  def log_weight():
  	socket_open(SERVER_IP,SERVER_PORT)
  	socket_send_string("LOG_WEIGHT")
  	sleep(0.5)
  	socket_close()
  end

  def send_target_info():
  	socket_open(SERVER_IP,SERVER_PORT)
  	socket_send_string("SET_TARGET:" + to_str(target_weight))
  	sleep(0.2)
  	socket_close()
  end
  def send_powder_info():
  	socket_open(SERVER_IP,SERVER_PORT)
  	socket_send_string("SET_POWDER:" + Pow_name)
  	sleep(0.2)
  	socket_close()
  end
  def send_spatula_info():
  	socket_open(SERVER_IP,SERVER_PORT)
  	socket_send_string("SET_SPATULA:" + spatula)
  	#sleep(1)

  	#local fl = socket_read_ascii_float(4)
    	#socket_close()

    	#global s_depth = fl[1]
    	#global s_length = fl[2]
   	#global s_volume = fl[3]
   	#global ry_theta  = fl[4]
  	sleep(0.2)

  end

  def send_level_info():
  	socket_open(SERVER_IP,SERVER_PORT)
  	socket_send_string("SET_LEVEL:" + to_str(level))
  	sleep(0.2)
  	socket_close()
  end

  def get_cont_weight():
    socket_open(SERVER_IP, SERVER_PORT)
    #rq_open_and_wait()
    cmd = "GET_CONT_WEIGHT"
    socket_send_string(cmd)
    sync()
    sleep(0.5)
    receiveFromSer = socket_read_ascii_float(1)
    socket_close()
    return receiveFromSer[1]
  end

  $ 22 "BeforeStarts"
  $ 23 "uLM"
  $ 24 "CMD_Stop≔ False "
  global CMD_Stop=  False
  $ 25 "CMD_Abort≔ False "
  global CMD_Abort=  False
  $ 26 "CMD_Clear≔ False "
  global CMD_Clear=  False
  $ 27 "STATE≔1"
  global STATE=1
  $ 28 "STATE_Info≔''"
  global STATE_Info=""
  $ 29 "ARM_Referenced≔ False "
  global ARM_Referenced=  False
  $ 30 "zero_ftsensor()"
  zero_ftsensor()
  $ 31 "poses init"
  $ 32 "PSE_A≔p[0,0,0,0,0,0]"
  global PSE_A=p[0,0,0,0,0,0]
  $ 33 "PSE_A_H≔p[0,0,0,0,0,0]"
  global PSE_A_H=p[0,0,0,0,0,0]
  $ 34 "PSE_R≔p[0,0,0,0,0,0]"
  global PSE_R=p[0,0,0,0,0,0]
  $ 35 "PSE_R_H≔p[0,0,0,0,0,0]"
  global PSE_R_H=p[0,0,0,0,0,0]
  $ 36 "PSE_T≔p[0,0,0,0,0,0]"
  global PSE_T=p[0,0,0,0,0,0]
  $ 37 "PSE_T_H≔p[0,0,0,0,0,0]"
  global PSE_T_H=p[0,0,0,0,0,0]
  $ 38 "PSE_C_E≔p[0,0,0,0,0,0]"
  global PSE_C_E=p[0,0,0,0,0,0]
  $ 39 "PSE_C_H≔p[0,0,0,0,0,0]"
  global PSE_C_H=p[0,0,0,0,0,0]
  $ 40 "PSE_C_S≔p[0,0,0,0,0,0]"
  global PSE_C_S=p[0,0,0,0,0,0]
  $ 41 "init_home_by_cartesian_pose(p[0,-0.400,0.300,0,0,0])"
  init_home_by_cartesian_pose(p[0,-0.400,0.300,0,0,0])
  $ 42 "Clearing"
  $ 43 "reset_error()"
  reset_error()
  $ 44 "reset_warning()"
  reset_warning()
  $ 45 "uGo"
  $ 47 "ugo_init( True ,'http://192.168.12.120:10001')"
  ugo_init(  True  ,"http://192.168.12.120:10001")
  $ 48 "ugo_update_outputs()"
  ugo_update_outputs()
  $ 49 "App"
  $ 50 "'ADD APPLICATION SPECIFIC COMMANDS'"
  # 'ADD APPLICATION SPECIFIC COMMANDS'
  $ 51 "Tools"
  $ 52 "OBJ_Picked≔gripper_has_object()"
  global OBJ_Picked=gripper_has_object()
  $ 53 "If OBJ_Picked"
  if (OBJ_Picked):
    # begin: URCap Program Node
    #   Source: Robotiq_Grippers, 3.17.0.105337, Robotiq Inc.
    #   Type: Gripper Activate
    $ 54 "Gripper Activate"

    kill rq_gripper_communication_thread
    rq_gripper_communication_thread_started = False
    rq_close_gripper_socket("1")
    rq_close_gripper_socket("2")
    rq_close_gripper_socket("3")
    rq_close_gripper_socket("4")

    rq_init_comm_if_connected(9, "1")
    rq_init_comm_if_connected(2, "2")
    rq_init_comm_if_connected(3, "3")
    rq_init_comm_if_connected(4, "4")
    rq_print_connected_grippers()
    rq_gripper_communication_thread = run rq_gripper_communication()

    while(not rq_gripper_communication_thread_started):
        sleep(0.008)
    end

    rq_set_max_current_for_all_grippers()

    reset_and_activate = False

    rq_activate_all_grippers(False)
    # end: URCap Program Node
  else:
    $ 55 "Else" "noBreak"
    # begin: URCap Program Node
    #   Source: Robotiq_Grippers, 3.17.0.105337, Robotiq Inc.
    #   Type: Gripper Activate
    $ 56 "Gripper Reset and Activate"

    kill rq_gripper_communication_thread
    rq_gripper_communication_thread_started = False
    rq_close_gripper_socket("1")
    rq_close_gripper_socket("2")
    rq_close_gripper_socket("3")
    rq_close_gripper_socket("4")

    rq_init_comm_if_connected(9, "1")
    rq_init_comm_if_connected(2, "2")
    rq_init_comm_if_connected(3, "3")
    rq_init_comm_if_connected(4, "4")
    rq_print_connected_grippers()
    rq_gripper_communication_thread = run rq_gripper_communication()

    while(not rq_gripper_communication_thread_started):
        sleep(0.008)
    end

    rq_set_max_current_for_all_grippers()

    reset_and_activate = True

    rq_activate_all_grippers(True)
    # end: URCap Program Node
  end
  $ 57 "zero_ftsensor()"
  zero_ftsensor()
  $ 58 "EXTT"
  $ 59 "Set GRP_3F_Enable=Off"
  set_standard_digital_out(4, False)
  $ 60 "Set BarcodeTrigger=Off"
  set_standard_digital_out(6, False)
  $ 61 "Set GRP_3F_Decap=Off"
  set_standard_digital_out(3, False)
  $ 62 "Set GRP_3F_Cap=Off"
  set_standard_digital_out(2, False)
  $ 63 "Set GRP_3F_Open=Off"
  set_standard_digital_out(5, False)
  $ 64 "PSE_T≔get_tool_free_pose(dir=[0,0,0.150], move_in_base_frame=True)"
  global PSE_T=get_tool_free_pose(dir=[0,0,0.150], move_in_base_frame=True)
  $ 65 "If is_reachable(Base_const, [PSE_T])"
  if (is_reachable(p[0.0,0.0,0.0,0.0,0.0,0.0], [PSE_T])):
    $ 66 "MoveL"
    $ 67 "PSE_T" "breakAfter"
    movel(PSE_T, a=1.2, v=0.15)
  end
  $ 68 "powder dispensing variable init"
  $ 69 "Start_thread≔ False "
  global Start_thread=  False
  $ 70 "vib_thread≔ False "
  global vib_thread=  False
  $ 71 "w_full_thread≔ False "
  global w_full_thread=  False
  $ 72 "d_cc≔0.07"
  global d_cc=0.07
  $ 73 "kp≔0.0035"
  global kp=0.0035
  $ 74 "ki≔0.0001"
  global ki=0.0001
  $ 75 "kd≔0.003"
  global kd=0.003
  $ 76 "dt≔0.2"
  global dt=0.2
  $ 77 "Integral_error≔0"
  global Integral_error=0
  $ 78 "current_error≔0"
  global current_error=0
  $ 79 "previous_error≔0"
  global previous_error=0
  $ 80 "tilt_increment≔0"
  global tilt_increment=0
  $ 81 "tilt_angle≔0"
  global tilt_angle=0
  $ 82 "diff≔0"
  global diff=0
  $ 83 "tilt_to_home()"
  tilt_to_home()
  $ 84 "switch_spat_M≔ True "
  global switch_spat_M=  True
  $ 85 "switch_spat_S≔ True "
  global switch_spat_S=  True
  $ 86 "switch_spat_F_M≔ True "
  global switch_spat_F_M=  True
  $ 87 "switch_spat_F_S≔ True "
  global switch_spat_F_S=  True
  $ 88 "last_scale≔0"
  global last_scale=0
  $ 817 "Thread_1"
  thread Thread_1():
    while (True):
      $ 818 "If Start_thread≟ True "
      if (Start_thread ==   True  ):
        $ 819 "weight_value≔get_weight()"
        global weight_value=get_weight()
        $ 820 "diff≔target_weight-weight_value"
        global diff=target_weight-weight_value
        $ 821 "Wait: 0.2"
        sleep(0.2)
        $ 822 "sync()"
        sync()
      end
      $ 823 "sync()"
      sync()
    end
  end
  threadId_Thread_1 = run Thread_1()
  $ 824 "Thread_2"
  thread Thread_2():
    while (True):
      $ 825 "Loop vib_thread≟ True "
      thread Thread_while_825():
        while (True):
          $ 826 "diff≔target_weight-weight_value"
          global diff=target_weight-weight_value
          $ 827 "If diff>0.02 and spatula≠'spatula_flat_S' "
          global thread_flag_827=0
          thread Thread_if_827():
            $ 829 "Set AO[0]=4.0"
            set_standard_analog_out(0, 0.4)
            thread_flag_827 = 1
          end
          if (diff>0.02  and  spatula != "spatula_flat_S" ):
            global thread_handler_827=run Thread_if_827()
            while (thread_flag_827 == 0):
              if not(diff>0.02  and  spatula != "spatula_flat_S" ):
                kill thread_handler_827
                thread_flag_827 = 2
              else:
                sync()
              end
            end
          else:
            thread_flag_827 = 2
          end
          if (thread_flag_827 == 2):
            $ 830 "ElseIf diff>0.02 and spatula≟'spatula_flat_S'"
            if (diff>0.02 and spatula == "spatula_flat_S"):
              $ 831 "vibration_3()"
              vibration_3()
            else:
              $ 832 "ElseIf diff≤0.03"
              global thread_flag_832=0
              thread Thread_if_832():
                $ 833 "vibration_2()"
                vibration_2()
                thread_flag_832 = 1
              end
              if (diff <= 0.03):
                global thread_handler_832=run Thread_if_832()
                while (thread_flag_832 == 0):
                  if not(diff <= 0.03):
                    kill thread_handler_832
                    thread_flag_832 = 2
                  else:
                    sync()
                  end
                end
              else:
                thread_flag_832 = 2
              end
              if (thread_flag_832 == 2):
                $ 834 "Else" "noBreak"
                $ 835 "Set AO[0]=0.0"
                set_standard_analog_out(0, 0.0)
              end
            end
          end
        end
      end
      if (vib_thread ==   True  ):
        global thread_handler_825=run Thread_while_825()
        while (vib_thread ==   True  ):
          sync()
        end
        kill thread_handler_825
      end
      $ 836 "sync()"
      sync()
    end
  end
  threadId_Thread_2 = run Thread_2()
  $ 837 "Thread_3"
  thread Thread_3():
    while (True):
      $ 838 "If w_full_thread≟ True "
      if (w_full_thread ==   True  ):
        $ 839 "aa_weight_cont≔get_cont_weight()"
        global aa_weight_cont=get_cont_weight()
        $ 840 "Wait: 0.2"
        sleep(0.2)
        $ 841 "sync()"
        sync()
      end
      $ 842 "sync()"
      sync()
    end
  end
  threadId_Thread_3 = run Thread_3()
  while (True):
    $ 89 "Robot Program"
    $ 90 "MAIN"
    $ 91 "command_manager(external_control='uGO', cond_suspend=(ITM_Manipulated and AMR_AtTarget and AMR_Charging and AMR_Battery<40), cond_unsuspend=(AMR_Battery≟60))"
    command_manager(external_control="uGO", cond_suspend=(ITM_Manipulated  and  AMR_AtTarget  and  AMR_Charging  and  AMR_Battery<40), cond_unsuspend=(AMR_Battery == 60))
    $ 92 "log_state(STATE_Info)"
    log_state(STATE_Info)
    $ 93 "Switch STATE"
    switch_1 = STATE
    $ 94 "Case 1"
    if (1 == switch_1):
      $ 95 "Stopping"
      $ 96 "STATE_Info≔'Stopping'"
      global STATE_Info="Stopping"
      $ 97 "end_freedrive_mode()"
      end_freedrive_mode()
      $ 98 "Set"
      set_tcp(p[0.0,0.0,0.161,3.1415,0.0,0.0])
      $ 99 "PSE_T≔get_tool_free_pose(dir=[0,0,0.150], move_in_base_frame=True)"
      global PSE_T=get_tool_free_pose(dir=[0,0,0.150], move_in_base_frame=True)
      $ 100 "If is_reachable(Base_const, [PSE_T])"
      if (is_reachable(p[0.0,0.0,0.0,0.0,0.0,0.0], [PSE_T])):
        $ 101 "MoveL"
        $ 102 "PSE_T" "breakAfter"
        movel(PSE_T, a=1.2, v=0.15)
      end
      $ 103 "do_transition(keep_rxry=OBJ_Picked, r=0)"
      do_transition(keep_rxry=OBJ_Picked, r=0)
      $ 112 "Call Sub_AMR_MiR_V3"
      Sub_AMR_MiR_V3()
      $ 113 "If stopping() and AMR_Done"
      if (stopping()  and  AMR_Done):
        $ 114 "STATE≔2"
        global STATE=2
        $ 115 "ugo_update_outputs()"
        ugo_update_outputs()
      end
    elif (2 == switch_1):
      $ 116 "Case 2"
      $ 117 "Stopped"
      $ 118 "STATE_Info≔'Stopped'"
      global STATE_Info="Stopped"
      $ 119 "Call Sub_AMR_MiR_V3"
      Sub_AMR_MiR_V3()
      $ 120 "If CMD_Reset  or PB_Start"
      if (CMD_Reset   or  get_standard_digital_in(0)):
        $ 121 "STATE≔3"
        global STATE=3
        $ 122 "ugo_update_outputs()"
        ugo_update_outputs()
      end
    elif (3 == switch_1):
      $ 123 "Case 3"
      $ 124 " Resetting"
      $ 125 "STATE_Info≔'Resetting'"
      global STATE_Info="Resetting"
      $ 126 "uML"
      $ 127 "reset_error()"
      reset_error()
      $ 128 "reset_warning()"
      reset_warning()
      $ 129 "PROCESS_Step≔0"
      global PROCESS_Step=0
      $ 130 "PROCESS_Info≔''"
      global PROCESS_Info=""
      $ 131 "ARM_Referenced≔ False "
      global ARM_Referenced=  False
      $ 132 "WRK_Done≔ False "
      global WRK_Done=  False
      $ 133 "ITM_Prepared≔ False "
      global ITM_Prepared=  False
      $ 134 "ITM_Manipulated≔ False "
      global ITM_Manipulated=  False
      $ 135 "STP≔0"
      global STP=0
      $ 136 "Action≔0"
      global Action=0
      $ 137 "Action_Info≔''"
      global Action_Info=""
      $ 138 "ITM_ID≔0"
      global ITM_ID=0
      $ 139 "JIG≔0"
      global JIG=0
      $ 140 "JIG_Slot≔0"
      global JIG_Slot=0
      $ 141 "Task_info≔''"
      global Task_info=""
      $ 142 "Set"
      set_tcp(p[0.0,0.0,0.161,3.1415,0.0,0.0])
      $ 143 "App"
      $ 144 "'ADD APPLICATION SPECIFIC COMMANDS'"
      # 'ADD APPLICATION SPECIFIC COMMANDS'
      $ 145 "OBJ_Type≔0"
      global OBJ_Type=0
      $ 146 "OBJ_Nbr≔0"
      global OBJ_Nbr=0
      $ 147 "If CNT_Rack_Output≥50"
      if (CNT_Rack_Output >= 50):
        $ 148 "CNT_Rack_Output≔0"
        global CNT_Rack_Output=0
      end
      $ 149 "TASK≔struct(ID=0, NAVI=struct(target=0, footprint=0, protectiveOff=0, dock=0), WORK=struct(ITM_ID_Src=0, JIG_ID_Src=0, OBJ_Nbr_Src=0, ACT_Src=0, ITM_ID_Tgt=0, JIG_ID_Tgt=0, OBJ_Nbr_Tgt=0, ACT_Tgt=0, OBJ_Type=0))"
      global TASK=struct(ID=0, NAVI=struct(target=0, footprint=0, protectiveOff=0, dock=0), WORK=struct(ITM_ID_Src=0, JIG_ID_Src=0, OBJ_Nbr_Src=0, ACT_Src=0, ITM_ID_Tgt=0, JIG_ID_Tgt=0, OBJ_Nbr_Tgt=0, ACT_Tgt=0, OBJ_Type=0))
      $ 150 "Call Sub_AMR_MiR_V3"
      Sub_AMR_MiR_V3()
      $ 151 "If resetting() and AMR_Done"
      if (resetting()  and  AMR_Done):
        $ 152 "STATE≔4"
        global STATE=4
        $ 153 "ugo_update_outputs()"
        ugo_update_outputs()
      end
    elif (4 == switch_1):
      $ 154 "Case 4"
      $ 155 "Idle"
      $ 156 "STATE_Info≔'Idle'"
      global STATE_Info="Idle"
      $ 157 "If CMD_Start"
      if (CMD_Start):
        $ 158 "STATE≔5"
        global STATE=5
        $ 159 "ugo_update_outputs()"
        ugo_update_outputs()
      end
    elif (5 == switch_1):
      $ 160 "Case 5"
      $ 161 "Starting"
      $ 162 "STATE_Info≔'Starting'"
      global STATE_Info="Starting"
      $ 163 "'ADD COMMANDS WHAT TO START WITH'"
      # 'ADD COMMANDS WHAT TO START WITH'
      $ 164 "Call Sub_AMR_MiR_V3"
      Sub_AMR_MiR_V3()
      $ 165 "get ugo data"
      $ 166 "Assign Tasks"
      $ 167 "TASK.ID = ugo_get_task()"
      TASK.ID = ugo_get_task()
      $ 168 "If TASK.ID≟1"
      if (TASK.ID == 1):
        $ 169 "Task_info≔'Charge'"
        global Task_info="Charge"
        $ 170 "Parameters"
        $ 171 "AMR_PosTarget≔1"
        global AMR_PosTarget=1
      else:
        $ 172 "ElseIf TASK.ID≟9"
        if (TASK.ID == 9):
          $ 173 "'Pick Sarstedt Rack from Variable source'"
          # 'Pick Sarstedt Rack from Variable source'
          $ 174 "Task_info≔'Navigate to Target'"
          global Task_info="Navigate to Target"
          $ 175 "Parameters"
          $ 176 "AMR_PosTarget≔UGO.read_input('00','ITM_ID')"
          global AMR_PosTarget=UGO.read_input("00","ITM_ID")
        else:
          $ 177 "ElseIf TASK.ID≟13"
          if (TASK.ID == 13):
            $ 178 "Task_info≔'Dose Powder'"
            global Task_info="Dose Powder"
            $ 179 "Parameters"
            $ 180 "ITM_ID≔1"
            global ITM_ID=1
            $ 181 "W_now≔(UGO.read_input('00','Container_weight'))/1000"
            global W_now=(UGO.read_input("00","Container_weight"))/1000
            $ 182 "Pow_name≔(UGO.read_input('00','Powder_name'))"
            global Pow_name=(UGO.read_input("00","Powder_name"))
            $ 183 "target_weight≔(UGO.read_input('00','Target_weight'))/1000"
            global target_weight=(UGO.read_input("00","Target_weight"))/1000
            $ 184 "send_picking_info(Pow_name,target_weight)"
            send_picking_info(Pow_name,target_weight)
            $ 185 "w_dosed_total≔0"
            global w_dosed_total=0
            $ 186 "OBJ_Type≔6"
            global OBJ_Type=6
            $ 187 "JIG≔17"
            global JIG=17
            $ 188 "AMR_PosTarget≔5"
            global AMR_PosTarget=5
          else:
            $ 189 "ElseIf TASK.ID≟49"
            if (TASK.ID == 49):
              $ 190 "Task_info≔'Pick Containers'"
              global Task_info="Pick Containers"
              $ 191 "Parameters"
              $ 192 "ITM_ID≔1"
              global ITM_ID=1
              $ 193 "OBJ_Type≔6"
              global OBJ_Type=6
              $ 194 "JIG≔15"
              global JIG=15
              $ 195 "AMR_PosTarget≔3"
              global AMR_PosTarget=3
            else:
              $ 196 "ElseIf TASK.ID≟50"
              if (TASK.ID == 50):
                $ 197 "Task_info≔'Decap Containers'"
                global Task_info="Decap Containers"
                $ 198 "Parameters"
                $ 199 "ITM_ID≔1"
                global ITM_ID=1
                $ 200 "OBJ_Type≔6"
                global OBJ_Type=6
                $ 201 "JIG≔16"
                global JIG=16
                $ 202 "AMR_PosTarget≔5"
                global AMR_PosTarget=5
              else:
                $ 203 "ElseIf TASK.ID≟51"
                if (TASK.ID == 51):
                  $ 204 "Task_info≔'Detect Spatula and transfer powder'"
                  global Task_info="Detect Spatula and transfer powder"
                  $ 205 "Parameters"
                  $ 206 "ITM_ID≔1"
                  global ITM_ID=1
                  $ 207 "target_weight≔(UGO.read_input('00','Target_weight'))/1000"
                  global target_weight=(UGO.read_input("00","Target_weight"))/1000
                  $ 208 "OBJ_Type≔8"
                  global OBJ_Type=8
                  $ 209 "JIG≔16"
                  global JIG=16
                  $ 210 "AMR_PosTarget≔5"
                  global AMR_PosTarget=5
                else:
                  $ 211 "ElseIf TASK.ID≟52"
                  if (TASK.ID == 52):
                    $ 212 "Task_info≔'Pick Powder'"
                    global Task_info="Pick Powder"
                    $ 213 "Parameters"
                    $ 214 "ITM_ID≔1"
                    global ITM_ID=1
                    $ 216 "OBJ_Type≔6"
                    global OBJ_Type=6
                    $ 217 "JIG≔15"
                    global JIG=15
                    $ 218 "AMR_PosTarget≔3"
                    global AMR_PosTarget=3
                  else:
                    $ 219 "ElseIf TASK.ID≟53"
                    if (TASK.ID == 53):
                      $ 220 "Task_info≔'Decap Powder'"
                      global Task_info="Decap Powder"
                      $ 221 "Parameters"
                      $ 222 "ITM_ID≔1"
                      global ITM_ID=1
                      $ 223 "OBJ_Type≔6"
                      global OBJ_Type=6
                      $ 224 "JIG≔1"
                      global JIG=1
                      $ 225 "AMR_PosTarget≔5"
                      global AMR_PosTarget=5
                    else:
                      $ 226 "ElseIf TASK.ID≟54"
                      if (TASK.ID == 54):
                        $ 227 "Task_info≔'Empty and swap Powder container'"
                        global Task_info="Empty and swap Powder container"
                        $ 236 "Parameters"
                        $ 237 "ITM_ID≔1"
                        global ITM_ID=1
                        $ 239 "W_now≔(UGO.read_input('00','Container_weight'))/1000"
                        global W_now=(UGO.read_input("00","Container_weight"))/1000
                        $ 240 "Pow_name≔(UGO.read_input('00','Powder_name'))"
                        global Pow_name=(UGO.read_input("00","Powder_name"))
                        $ 243 "OBJ_Type≔6"
                        global OBJ_Type=6
                        $ 244 "JIG≔17"
                        global JIG=17
                        $ 245 "AMR_PosTarget≔5"
                        global AMR_PosTarget=5
                      else:
                        $ 246 "ElseIf TASK.ID≟55"
                        if (TASK.ID == 55):
                          $ 247 "Task_info≔'Place Powder'"
                          global Task_info="Place Powder"
                          $ 248 "Parameters"
                          $ 249 "ITM_ID≔1"
                          global ITM_ID=1
                          $ 250 "OBJ_Type≔6"
                          global OBJ_Type=6
                          $ 251 "JIG≔21"
                          global JIG=21
                          $ 252 "AMR_PosTarget≔5"
                          global AMR_PosTarget=5
                        else:
                          $ 253 "ElseIf TASK.ID≟56"
                          if (TASK.ID == 56):
                            $ 254 "Task_info≔'Dose Powder'"
                            global Task_info="Dose Powder"
                            $ 255 "Parameters"
                            $ 256 "ITM_ID≔1"
                            global ITM_ID=1
                            $ 257 "target_weight≔(UGO.read_input('00','Target_weight'))/1000"
                            global target_weight=(UGO.read_input("00","Target_weight"))/1000
                            $ 258 "W_now≔(UGO.read_input('00','Container_weight'))/1000"
                            global W_now=(UGO.read_input("00","Container_weight"))/1000
                            $ 259 "Pow_name≔(UGO.read_input('00','Powder_name'))"
                            global Pow_name=(UGO.read_input("00","Powder_name"))
                            $ 260 "OBJ_Type≔6"
                            global OBJ_Type=6
                            $ 261 "JIG≔17"
                            global JIG=17
                            $ 262 "AMR_PosTarget≔5"
                            global AMR_PosTarget=5
                          else:
                            $ 263 "ElseIf TASK.ID≟57"
                            if (TASK.ID == 57):
                              $ 264 "Task_info≔'Recipe Powder dosing'"
                              global Task_info="Recipe Powder dosing"
                              $ 265 "Parameters"
                              $ 266 "ITM_ID≔1"
                              global ITM_ID=1
                              $ 267 "Pow_A≔(UGO.read_input('00','PowderA'))"
                              global Pow_A=(UGO.read_input("00","PowderA"))
                              $ 268 "Pow_B≔(UGO.read_input('00','PowderB'))"
                              global Pow_B=(UGO.read_input("00","PowderB"))
                              $ 269 "Pow_C≔(UGO.read_input('00','PowderC'))"
                              global Pow_C=(UGO.read_input("00","PowderC"))
                              $ 270 "Total_weight≔(UGO.read_input('00','Total_weight'))/1000"
                              global Total_weight=(UGO.read_input("00","Total_weight"))/1000
                              $ 271 "Pow_A_percent≔(UGO.read_input('00','PowderA_percentage'))/100"
                              global Pow_A_percent=(UGO.read_input("00","PowderA_percentage"))/100
                              $ 272 "Pow_B_percent≔(UGO.read_input('00','PowderB_percentage'))/100"
                              global Pow_B_percent=(UGO.read_input("00","PowderB_percentage"))/100
                              $ 273 "Pow_C_percent≔(UGO.read_input('00','PowderC_percentage'))/100"
                              global Pow_C_percent=(UGO.read_input("00","PowderC_percentage"))/100
                              $ 274 "OBJ_Type≔6"
                              global OBJ_Type=6
                              $ 275 "JIG≔17"
                              global JIG=17
                              $ 276 "AMR_PosTarget≔5"
                              global AMR_PosTarget=5
                            else:
                              $ 277 "ElseIf TASK.ID≟58"
                              if (TASK.ID == 58):
                                $ 278 "Task_info≔'Pick Powder containers'"
                                global Task_info="Pick Powder containers"
                                $ 279 "Parameters"
                                $ 280 "ITM_ID≔1"
                                global ITM_ID=1
                                $ 281 "OBJ_Type≔6"
                                global OBJ_Type=6
                                $ 282 "JIG≔15"
                                global JIG=15
                                $ 283 "AMR_PosTarget≔3"
                                global AMR_PosTarget=3
                              else:
                                $ 284 "ElseIf TASK.ID≟59"
                                if (TASK.ID == 59):
                                  $ 285 "Task_info≔'Empty Powder container'"
                                  global Task_info="Empty Powder container"
                                  $ 286 "Parameters"
                                  $ 287 "ITM_ID≔1"
                                  global ITM_ID=1
                                  $ 289 "Pow_name≔(UGO.read_input('00','Powder_name'))"
                                  global Pow_name=(UGO.read_input("00","Powder_name"))
                                  $ 291 "target_weight≔aa_weight_cont-empty_weight_g"
                                  global target_weight=aa_weight_cont-empty_weight_g
                                  $ 292 "send_picking_info(Pow_name,target_weight)"
                                  send_picking_info(Pow_name,target_weight)
                                  $ 293 "w_dosed_total≔0"
                                  global w_dosed_total=0
                                  $ 294 "OBJ_Type≔6"
                                  global OBJ_Type=6
                                  $ 295 "JIG≔17"
                                  global JIG=17
                                  $ 296 "AMR_PosTarget≔5"
                                  global AMR_PosTarget=5
                                else:
                                  $ 297 "ElseIf TASK.ID≟61"
                                  if (TASK.ID == 61):
                                    $ 298 "Task_info≔'Weigh, Place & Decap'"
                                    global Task_info="Weigh, Place & Decap"
                                    $ 299 "Parameters"
                                    $ 300 "ITM_ID≔1"
                                    global ITM_ID=1
                                    $ 301 "OBJ_Type≔6"
                                    global OBJ_Type=6
                                    $ 302 "JIG≔21"
                                    global JIG=21
                                    $ 303 "AMR_PosTarget≔5"
                                    global AMR_PosTarget=5
                                  else:
                                    $ 304 "Else" "noBreak"
                                    $ 305 "set_error(ERROR_WRONG_ORDER)"
                                    set_error(ERROR_WRONG_ORDER)
                                  end
                                end
                              end
                            end
                          end
                        end
                      end
                    end
                  end
                end
              end
            end
          end
        end
      end
      $ 306 "test ugo"
      $ 307 "Wait: 0.2"
      sleep(0.2)
      $ 308 "ugo_update_outputs()"
      ugo_update_outputs()
      $ 309 "If starting() and AMR_Done"
      if (starting()  and  AMR_Done):
        $ 310 "log_message(Task_info, 'New Task: ')"
        log_message(Task_info, "New Task: ")
        $ 311 "log_message(to_str(TASK.ID), 'Task_ID: ')"
        log_message(to_str(TASK.ID), "Task_ID: ")
        $ 312 "do_transition(keep_rxry=OBJ_Picked)"
        do_transition(keep_rxry=OBJ_Picked)
        $ 313 "STATE≔6"
        global STATE=6
        $ 314 "ugo_update_outputs()"
        ugo_update_outputs()
      end
    elif (6 == switch_1):
      $ 315 "Case 6"
      $ 316 "Execute"
      $ 317 "STATE_Info≔'Execute'"
      global STATE_Info="Execute"
      $ 318 "If  not CMD_Hold and not CMD_Suspend"
      global thread_flag_318=0
      thread Thread_if_318():
        $ 319 "Switch PROCESS_Step"
        switch_2 = PROCESS_Step
        $ 320 "Case 0"
        if (0 == switch_2):
          $ 321 "PROCESS_Info≔'process control'"
          global PROCESS_Info="process control"
          $ 322 "log_process(PROCESS_Info)"
          log_process(PROCESS_Info)
          $ 323 "process control"
          $ 324 "If  not AMR_AtTarget"
          if (  not  AMR_AtTarget):
            $ 325 "PROCESS_Step≔1"
            global PROCESS_Step=1
          else:
            $ 326 "ElseIf (( not ITM_Prepared and  not WRK_Done) or (ITM_Prepared and WRK_Done))"
            if (((  not  ITM_Prepared  and    not  WRK_Done)  or  (ITM_Prepared  and  WRK_Done))):
              $ 327 "PROCESS_Step≔2"
              global PROCESS_Step=2
            else:
              $ 328 "ElseIf  not WRK_Done"
              if (  not  WRK_Done):
                $ 329 "PROCESS_Step≔3"
                global PROCESS_Step=3
              else:
                $ 330 "Else" "noBreak"
                $ 331 "task finished"
                $ 332 "PROCESS_Info≔''"
                global PROCESS_Info=""
                $ 333 "STATE≔7"
                global STATE=7
                $ 334 "ugo_update_outputs()"
                ugo_update_outputs()
              end
            end
          end
        elif (1 == switch_2):
          $ 335 "Case 1"
          $ 336 "navigate"
          $ 337 "'MOVING THE uML'"
          # 'MOVING THE uML'
          $ 338 "PROCESS_Info≔'move to target'"
          global PROCESS_Info="move to target"
          $ 339 "log_process(PROCESS_Info)"
          log_process(PROCESS_Info)
          $ 340 "If TASK.ID≟1"
          if (TASK.ID == 1):
            $ 341 "Action≔51"
            global Action=51
          else:
            $ 342 "Else" "noBreak"
            $ 343 "Action≔52"
            global Action=52
          end
          $ 344 "Call Sub_AMR_MiR_V3"
          Sub_AMR_MiR_V3()
          $ 345 "If AMR_Done"
          if (AMR_Done):
            $ 346 "PROCESS_Step≔0"
            global PROCESS_Step=0
          end
        elif (2 == switch_2):
          $ 347 "Case 2"
          $ 348 "prepare"
          $ 349 "'THINGS THAT HAVE TO BE DONE ONCE IN A SEQUENCE,WORKFLOW'"
          # 'THINGS THAT HAVE TO BE DONE ONCE IN A SEQUENCE,WORKFLOW'
          $ 350 "PROCESS_Info≔'prepare for work'"
          global PROCESS_Info="prepare for work"
          $ 351 "log_process(PROCESS_Info)"
          log_process(PROCESS_Info)
          $ 352 "If TASK.WORK.ITM_ID_Src>1"
          if (TASK.WORK.ITM_ID_Src>1):
            $ 353 "ITM_ID≔TASK.WORK.ITM_ID_Src"
            global ITM_ID=TASK.WORK.ITM_ID_Src
          else:
            $ 354 "ElseIf TASK.WORK.ITM_ID_Tgt>1"
            if (TASK.WORK.ITM_ID_Tgt>1):
              $ 355 "ITM_ID≔TASK.WORK.ITM_ID_Tgt"
              global ITM_ID=TASK.WORK.ITM_ID_Tgt
            end
          end
          $ 356 "If  not ARM_Referenced and (ITM_ID≠0)"
          if (  not  ARM_Referenced  and  (ITM_ID != 0)):
            $ 357 "STP≔1"
            global STP=1
          else:
            $ 358 "ElseIf ARM_Referenced or (ITM_ID≟0)"
            if (ARM_Referenced  or  (ITM_ID == 0)):
              $ 359 "STP≔2"
              global STP=2
            end
          end
          $ 360 "Switch STP"
          switch_3 = STP
          $ 361 "Case 1"
          if (1 == switch_3):
            $ 362 "reference"
            $ 363 "STP_Info≔'reference at target position'"
            global STP_Info="reference at target position"
            $ 364 "log_step(STP_Info)"
            log_step(STP_Info)
            $ 365 "If ITM_ID≟1"
            if (ITM_ID == 1):
              $ 366 "CAM_Done≔ True "
              global CAM_Done=  True
            else:
              $ 367 "Else" "noBreak"
              $ 368 "Action≔131"
              global Action=131
              $ 369 "Call Sub_Vision_V18"
              Sub_Vision_V18()
            end
            $ 371 "If CAM_Done and  not ERROR.FLAG"
            if (CAM_Done  and    not  ERROR.FLAG):
              $ 372 "log_step('ARM referenced')"
              log_step("ARM referenced")
              $ 373 "ARM_Referenced≔ True "
              global ARM_Referenced=  True
            end
          elif (2 == switch_3):
            $ 374 "Case 2"
            $ 375 "manipulate"
            $ 376 "STP_Info≔'manipulate item'"
            global STP_Info="manipulate item"
            $ 377 "log_step(STP_Info)"
            log_step(STP_Info)
            $ 378 "'In case pressing button is needed'"
            # 'In case pressing button is needed'
            $ 379 "If found_in_list(ITM_ID, ITM_ID_List)"
            if (found_in_list(ITM_ID, ITM_ID_List)):
              $ 380 "Switch ITM_ID"
              switch_4 = ITM_ID
              $ 381 "Case 0"
              if (0 == switch_4):
                $ 382 "ITM_Manipulated≔ not ITM_Manipulated"
                global ITM_Manipulated=  not  ITM_Manipulated
              elif (1 == switch_4):
                $ 383 "Case 1"
                $ 384 "ITM_Manipulated≔ not ITM_Manipulated"
                global ITM_Manipulated=  not  ITM_Manipulated
              elif (2 == switch_4):
                $ 385 "Case 2"
              else:
                $ 395 "Default Case"
                $ 396 "ITM_Manipulated≔ not ITM_Manipulated"
                global ITM_Manipulated=  not  ITM_Manipulated
              end
            end
          end
          $ 397 "ITM_Prepared≔(ITM_Manipulated or  not found_in_list(ITM_ID, ITM_ID_List)) and (ARM_Referenced or ITM_ID≟0) and  not WRK_Done"
          global ITM_Prepared=(ITM_Manipulated  or    not  found_in_list(ITM_ID, ITM_ID_List))  and  (ARM_Referenced  or  ITM_ID == 0)  and    not  WRK_Done
          $ 398 "STP≔0"
          global STP=0
          $ 399 "STP_Info≔''"
          global STP_Info=""
          $ 400 "PROCESS_Step≔0"
          global PROCESS_Step=0
        elif (3 == switch_2):
          $ 401 "Case 3"
          $ 402 "work"
          $ 403 "'ADD EVERY MACHINE, OBJECT, STATION TO WORK ON'"
          # 'ADD EVERY MACHINE, OBJECT, STATION TO WORK ON'
          $ 404 "Switch ITM_ID"
          switch_3 = ITM_ID
          $ 405 "Case 1"
          if (1 == switch_3):
            $ 406 "uLM"
            $ 407 "If TASK.ID≟12"
            if (TASK.ID == 12):
              $ 408 "fill racks"
              $ 409 "Action≔151"
              global Action=151
              $ 410 "Call Sub_Vision_V18"
              Sub_Vision_V18()
              $ 411 "If  not ERROR.FLAG"
              if (  not  ERROR.FLAG):
                $ 412 "Actions for the task"
                $ 413 "Action≔1"
                global Action=1
                $ 414 "JIG≔2"
                global JIG=2
                $ 415 "JIG_Slot≔CAM_Result[0]"
                global JIG_Slot=CAM_Result[0]
                $ 416 "OBJ_Nbr≔CAM_Result[0]"
                global OBJ_Nbr=CAM_Result[0]
                $ 417 "OBJ_Type≔2"
                global OBJ_Type=2
                $ 418 "Call Sub_Action_V4"
                Sub_Action_V4()
                $ 419 "If OBJ_Picked"
                if (OBJ_Picked):
                  $ 420 "CAM_Result.remove(0)"
                  CAM_Result.remove(0)
                  $ 421 "PRC_TubCounter≔PRC_TubCounter+1"
                  global PRC_TubCounter=PRC_TubCounter+1
                  $ 422 "If PRC_TubCounter%4≟0"
                  if (PRC_TubCounter%4 == 0):
                    $ 423 "JIG_Slot≔4"
                    global JIG_Slot=4
                  else:
                    $ 424 "Else" "noBreak"
                    $ 425 "JIG_Slot≔PRC_TubCounter%4"
                    global JIG_Slot=PRC_TubCounter%4
                  end
                  $ 426 "OBJ_Nbr≔ceil(PRC_TubCounter/4)"
                  global OBJ_Nbr=ceil(PRC_TubCounter/4)
                  $ 427 "Action≔2"
                  global Action=2
                  $ 428 "JIG≔4"
                  global JIG=4
                  $ 429 "Call Sub_Action_V4"
                  Sub_Action_V4()
                  $ 430 "Action≔151"
                  global Action=151
                  $ 431 "Call Sub_Vision_V18"
                  Sub_Vision_V18()
                end
              end
              $ 432 "If (CAM_Captures≥CAM_PRM_Retries) or (PRC_TubCounter≥32)"
              if ((CAM_Captures >= CAM_PRM_Retries)  or  (PRC_TubCounter >= 32)):
                $ 433 "PROCESS_Step≔0"
                global PROCESS_Step=0
                $ 434 "WRK_Done≔ True "
                global WRK_Done=  True
              end
            else:
              $ 435 "ElseIf TASK.ID≟13"
              if (TASK.ID == 13):
                $ 436 "Dose Powder"
                $ 437 "Action≔131"
                global Action=131
                $ 438 "Call Sub_Vision_V18"
                Sub_Vision_V18()
                $ 439 "Action≔34"
                global Action=34
                $ 440 "Call Sub_Action_V4"
                Sub_Action_V4()
                $ 441 "PROCESS_Step≔0"
                global PROCESS_Step=0
                $ 442 "WRK_Done≔ True "
                global WRK_Done=  True
              else:
                $ 443 "ElseIf TASK.ID≟49"
                if (TASK.ID == 49):
                  $ 444 "Pick Powder container"
                  $ 445 "Action≔131"
                  global Action=131
                  $ 446 "Call Sub_Vision_V18"
                  Sub_Vision_V18()
                  $ 447 "Action≔35"
                  global Action=35
                  $ 448 "Call Sub_Action_V4"
                  Sub_Action_V4()
                  $ 449 "PROCESS_Step≔0"
                  global PROCESS_Step=0
                  $ 450 "WRK_Done≔ True "
                  global WRK_Done=  True
                else:
                  $ 451 "ElseIf TASK.ID≟50"
                  if (TASK.ID == 50):
                    $ 452 "Decap containers"
                    $ 453 "Action≔36"
                    global Action=36
                    $ 454 "Call Sub_Action_V4"
                    Sub_Action_V4()
                    $ 455 "PROCESS_Step≔0"
                    global PROCESS_Step=0
                    $ 456 "WRK_Done≔ True "
                    global WRK_Done=  True
                  else:
                    $ 457 "ElseIf TASK.ID≟51"
                    if (TASK.ID == 51):
                      $ 458 "Detect Spatula and transfer powder"
                      $ 459 "Action≔131"
                      global Action=131
                      $ 460 "Call Sub_Vision_V18"
                      Sub_Vision_V18()
                      $ 461 "Action≔37"
                      global Action=37
                      $ 462 "Call Sub_Action_V4"
                      Sub_Action_V4()
                      $ 463 "PROCESS_Step≔0"
                      global PROCESS_Step=0
                      $ 464 "WRK_Done≔ True "
                      global WRK_Done=  True
                    else:
                      $ 465 "ElseIf TASK.ID≟52"
                      if (TASK.ID == 52):
                        $ 466 "Pick Powder container"
                        $ 467 "Action≔131"
                        global Action=131
                        $ 468 "Call Sub_Vision_V18"
                        Sub_Vision_V18()
                        $ 469 "Action≔39"
                        global Action=39
                        $ 470 "Call Sub_Action_V4"
                        Sub_Action_V4()
                        $ 471 "PROCESS_Step≔0"
                        global PROCESS_Step=0
                        $ 472 "WRK_Done≔ True "
                        global WRK_Done=  True
                      else:
                        $ 473 "ElseIf TASK.ID≟53"
                        if (TASK.ID == 53):
                          $ 474 "Decap containerA"
                          $ 475 "Action≔40"
                          global Action=40
                          $ 476 "Call Sub_Action_V4"
                          Sub_Action_V4()
                          $ 477 "PROCESS_Step≔0"
                          global PROCESS_Step=0
                          $ 478 "WRK_Done≔ True "
                          global WRK_Done=  True
                        else:
                          $ 479 "ElseIf TASK.ID≟55"
                          if (TASK.ID == 55):
                            $ 480 "Place Powder"
                            $ 481 "Action≔131"
                            global Action=131
                            $ 482 "Call Sub_Vision_V18"
                            Sub_Vision_V18()
                            $ 483 "Action≔41"
                            global Action=41
                            $ 484 "Call Sub_Action_V4"
                            Sub_Action_V4()
                            $ 485 "PROCESS_Step≔0"
                            global PROCESS_Step=0
                            $ 486 "WRK_Done≔ True "
                            global WRK_Done=  True
                          else:
                            $ 487 "ElseIf TASK.ID≟54"
                            if (TASK.ID == 54):
                              $ 488 "Empty and swap container"
                              $ 489 "Action≔131"
                              global Action=131
                              $ 490 "Call Sub_Vision_V18"
                              Sub_Vision_V18()
                              $ 491 "Action≔42"
                              global Action=42
                              $ 492 "Call Sub_Action_V4"
                              Sub_Action_V4()
                              $ 493 "PROCESS_Step≔0"
                              global PROCESS_Step=0
                              $ 494 "WRK_Done≔ True "
                              global WRK_Done=  True
                            else:
                              $ 495 "ElseIf TASK.ID≟56"
                              if (TASK.ID == 56):
                                $ 496 "Dispense Powder"
                                $ 497 "Action≔131"
                                global Action=131
                                $ 498 "Call Sub_Vision_V18"
                                Sub_Vision_V18()
                                $ 499 "Action≔43"
                                global Action=43
                                $ 500 "Call Sub_Action_V4"
                                Sub_Action_V4()
                                $ 501 "PROCESS_Step≔0"
                                global PROCESS_Step=0
                                $ 502 "WRK_Done≔ True "
                                global WRK_Done=  True
                              else:
                                $ 503 "ElseIf TASK.ID≟57"
                                if (TASK.ID == 57):
                                  $ 504 "Recipe Dosing"
                                  $ 505 "Action≔48"
                                  global Action=48
                                  $ 506 "Call Sub_Action_V4"
                                  Sub_Action_V4()
                                  $ 523 "PROCESS_Step≔0"
                                  global PROCESS_Step=0
                                  $ 524 "WRK_Done≔ True "
                                  global WRK_Done=  True
                                else:
                                  $ 525 "ElseIf TASK.ID≟58"
                                  if (TASK.ID == 58):
                                    $ 526 "Pick Powder containers"
                                    $ 527 "Num_cont_picked≔0"
                                    global Num_cont_picked=0
                                    $ 528 "powder_position≔'Position1'"
                                    global powder_position="Position1"
                                    $ 529 "Loop Num_cont_picked<3"
                                    while (Num_cont_picked<3):
                                      $ 530 "Action≔131"
                                      global Action=131
                                      $ 531 "Call Sub_Vision_V18"
                                      Sub_Vision_V18()
                                      $ 532 "Action≔47"
                                      global Action=47
                                      $ 533 "Call Sub_Action_V4"
                                      Sub_Action_V4()
                                    end
                                    $ 534 "PROCESS_Step≔0"
                                    global PROCESS_Step=0
                                    $ 535 "WRK_Done≔ True "
                                    global WRK_Done=  True
                                  else:
                                    $ 536 "ElseIf TASK.ID≟59"
                                    if (TASK.ID == 59):
                                      $ 537 "Empty powder container"
                                      $ 538 "Action≔131"
                                      global Action=131
                                      $ 539 "Call Sub_Vision_V18"
                                      Sub_Vision_V18()
                                      $ 540 "Action≔50"
                                      global Action=50
                                      $ 541 "Call Sub_Action_V4"
                                      Sub_Action_V4()
                                      $ 542 "PROCESS_Step≔0"
                                      global PROCESS_Step=0
                                      $ 543 "WRK_Done≔ True "
                                      global WRK_Done=  True
                                    else:
                                      $ 544 "ElseIf TASK.ID≟61"
                                      if (TASK.ID == 61):
                                        $ 545 "Place Powder"
                                        $ 546 "Action≔131"
                                        global Action=131
                                        $ 547 "Call Sub_Vision_V18"
                                        Sub_Vision_V18()
                                        $ 548 "Action≔51"
                                        global Action=51
                                        $ 549 "Call Sub_Action_V4"
                                        Sub_Action_V4()
                                        $ 550 "PROCESS_Step≔0"
                                        global PROCESS_Step=0
                                        $ 551 "WRK_Done≔ True "
                                        global WRK_Done=  True
                                      end
                                    end
                                  end
                                end
                              end
                            end
                          end
                        end
                      end
                    end
                  end
                end
              end
            end
          elif (2 == switch_3):
            $ 552 "Case 2"
          elif (5 == switch_3):
            $ 594 "Case 5"
          elif (20 == switch_3):
            $ 602 "Case 20"
          elif (43 == switch_3):
            $ 664 "Case 43"
          else:
            $ 672 "Default Case"
            $ 673 "WRK_Done≔ True "
            global WRK_Done=  True
            $ 674 "PROCESS_Step≔0"
            global PROCESS_Step=0
          end
        end
        thread_flag_318 = 1
      end
      if (  not  CMD_Hold and not CMD_Suspend):
        global thread_handler_318=run Thread_if_318()
        while (thread_flag_318 == 0):
          if not(  not  CMD_Hold and not CMD_Suspend):
            kill thread_handler_318
            thread_flag_318 = 2
          else:
            sync()
          end
        end
      else:
        thread_flag_318 = 2
      end
      $ 675 "If CMD_Hold"
      if (CMD_Hold):
        $ 676 "STATE≔9"
        global STATE=9
        $ 677 "ugo_update_outputs()"
        ugo_update_outputs()
      else:
        $ 678 "ElseIf CMD_Suspend"
        if (CMD_Suspend):
          $ 679 "STATE≔12"
          global STATE=12
          $ 680 "ugo_update_outputs()"
          ugo_update_outputs()
        end
      end
    elif (7 == switch_1):
      $ 681 "Case 7"
      $ 682 "Completing"
      $ 683 "STATE_Info≔'Completing'"
      global STATE_Info="Completing"
      $ 684 "'ADD COMMANDS FOR COMPLETING THE PROCESS'"
      # 'ADD COMMANDS FOR COMPLETING THE PROCESS'
      $ 685 "do_transition(keep_rxry=OBJ_Picked)"
      do_transition(keep_rxry=OBJ_Picked)
      $ 686 "Call Sub_AMR_MiR_V3"
      Sub_AMR_MiR_V3()
      $ 687 "If completing() and AMR_Done"
      if (completing()  and  AMR_Done):
        $ 688 "STATE≔8"
        global STATE=8
        $ 689 "ugo_update_outputs()"
        ugo_update_outputs()
      end
    elif (8 == switch_1):
      $ 690 "Case 8"
      $ 691 "Complete"
      $ 692 "STATE_Info≔'Complete'"
      global STATE_Info="Complete"
      $ 693 "If CMD_Reset"
      if (CMD_Reset):
        $ 694 "STATE≔3"
        global STATE=3
        $ 695 "ugo_update_outputs()"
        ugo_update_outputs()
      end
    elif (9 == switch_1):
      $ 696 "Case 9"
      $ 697 "Holding"
      $ 698 "STATE_Info≔'Holding'"
      global STATE_Info="Holding"
      $ 699 "stopl(0.5)"
      stopl(0.5)
      $ 700 "Call Sub_AMR_MiR_V3"
      Sub_AMR_MiR_V3()
      $ 701 "If holding() and AMR_Done"
      if (holding()  and  AMR_Done):
        $ 702 "STATE≔10"
        global STATE=10
        $ 703 "ugo_update_outputs()"
        ugo_update_outputs()
      end
    elif (10 == switch_1):
      $ 704 "Case 10"
      $ 705 "Held"
      $ 706 "STATE_Info≔'Held'"
      global STATE_Info="Held"
      $ 707 "If CMD_Unhold"
      if (CMD_Unhold):
        $ 708 "end_freedrive_mode()"
        end_freedrive_mode()
        $ 709 "STATE≔11"
        global STATE=11
        $ 710 "ugo_update_outputs()"
        ugo_update_outputs()
      else:
        $ 711 "ElseIf FNC_Freedrive"
        if (FNC_Freedrive):
          $ 712 "freedrive_mode()"
          freedrive_mode()
        else:
          $ 713 "Else" "noBreak"
          $ 714 "end_freedrive_mode()"
          end_freedrive_mode()
        end
      end
    elif (11 == switch_1):
      $ 715 "Case 11"
      $ 716 "Unholding"
      $ 717 "STATE_Info≔'Unholding'"
      global STATE_Info="Unholding"
      $ 718 "Clearing"
      $ 719 "Switch ERROR.ID"
      switch_2 = ERROR.ID
      $ 720 "Case 1002"
      if (1002 == switch_2):
        $ 721 "AMR_AtTarget≔ False "
        global AMR_AtTarget=  False
        $ 722 "ARM_Referenced≔ False "
        global ARM_Referenced=  False
        $ 723 "ITM_Prepared≔ False "
        global ITM_Prepared=  False
        $ 724 "PROCESS_Step≔1"
        global PROCESS_Step=1
      elif (2007 == switch_2):
        $ 725 "Case 2007"
        $ 726 "PROCESS_Step≔1"
        global PROCESS_Step=1
      end
      $ 727 "reset_error()"
      reset_error()
      $ 728 "reset_warning()"
      reset_warning()
      $ 729 "OBJ_Picked≔gripper_has_object()"
      global OBJ_Picked=gripper_has_object()
      $ 730 "Call Sub_AMR_MiR_V3"
      Sub_AMR_MiR_V3()
      $ 731 "If unholding() and AMR_Done"
      if (unholding()  and  AMR_Done):
        $ 732 "STATE≔6"
        global STATE=6
        $ 733 "ugo_update_outputs()"
        ugo_update_outputs()
      end
    elif (12 == switch_1):
      $ 734 "Case 12"
      $ 735 "Suspending"
      $ 736 "STATE_Info≔'Suspending'"
      global STATE_Info="Suspending"
      $ 737 "PROCESS_Info≔str_cat(PROCESS_Info, ' suspended')"
      global PROCESS_Info=str_cat(PROCESS_Info, " suspended")
      $ 738 "If suspending()"
      if (suspending()):
        $ 739 "STATE≔13"
        global STATE=13
        $ 740 "ugo_update_outputs()"
        ugo_update_outputs()
      end
    elif (13 == switch_1):
      $ 741 "Case 13"
      $ 742 "Suspended"
      $ 743 "STATE_Info≔'Suspended'"
      global STATE_Info="Suspended"
      $ 744 "Call Sub_AMR_MiR_V3"
      Sub_AMR_MiR_V3()
      $ 745 "If CMD_Unsuspend"
      if (CMD_Unsuspend):
        $ 746 "STATE≔14"
        global STATE=14
        $ 747 "ugo_update_outputs()"
        ugo_update_outputs()
      end
    elif (14 == switch_1):
      $ 748 "Case 14"
      $ 749 "Unsuspending"
      $ 750 "STATE_Info≔'Unsuspending'"
      global STATE_Info="Unsuspending"
      $ 751 "PROCESS_Step≔0"
      global PROCESS_Step=0
      $ 752 "If unsuspending()"
      if (unsuspending()):
        $ 753 "STATE≔6"
        global STATE=6
        $ 754 "ugo_update_outputs()"
        ugo_update_outputs()
      end
    elif (15 == switch_1):
      $ 755 "Case 15"
      $ 756 "Aborting"
      $ 757 "STATE_Info≔'Aborting'"
      global STATE_Info="Aborting"
      $ 758 "If aborting()"
      if (aborting()):
        $ 759 "STATE≔16"
        global STATE=16
        $ 760 "ugo_update_outputs()"
        ugo_update_outputs()
      end
    elif (16 == switch_1):
      $ 761 "Case 16"
      $ 762 "Aborted"
      $ 763 "STATE_Info≔'Aborted'"
      global STATE_Info="Aborted"
      $ 764 "If CMD_Clear"
      if (CMD_Clear):
        $ 765 "STATE≔17"
        global STATE=17
        $ 766 "ugo_update_outputs()"
        ugo_update_outputs()
      end
    elif (17 == switch_1):
      $ 767 "Case 17"
      $ 768 "Clearing"
      $ 769 "STATE_Info≔'Clearing'"
      global STATE_Info="Clearing"
      $ 770 "Clearing"
      $ 771 "reset_warning()"
      reset_warning()
      $ 772 "reset_error()"
      reset_error()
      $ 773 "If clearing()"
      if (clearing()):
        $ 774 "STATE≔2"
        global STATE=2
        $ 775 "ugo_update_outputs()"
        ugo_update_outputs()
      end
    end
    $ 776 "log_state(STATE_Info)"
    log_state(STATE_Info)
    $ 777 "log_warning(WARNING.MSG)"
    log_warning(WARNING.MSG)
    $ 778 "log_error(ERROR.MSG)"
    log_error(ERROR.MSG)
    $ 779 "Times"
    $ 780 "Switch STATE"
    switch_1 = STATE
    $ 781 "Case 1"
    if (1 == switch_1):
      $ 782 "TM_St_Stopping≔get_time(STATE_Times[STATE-1])"
      global TM_St_Stopping=get_time(STATE_Times[STATE-1])
    elif (2 == switch_1):
      $ 783 "Case 2"
      $ 784 "TM_St_Stopped≔get_time(STATE_Times[STATE-1])"
      global TM_St_Stopped=get_time(STATE_Times[STATE-1])
    elif (3 == switch_1):
      $ 785 "Case 3"
      $ 786 "TM_St_Resetting≔get_time(STATE_Times[STATE-1])"
      global TM_St_Resetting=get_time(STATE_Times[STATE-1])
    elif (4 == switch_1):
      $ 787 "Case 4"
      $ 788 "TM_St_Idle≔get_time(STATE_Times[STATE-1])"
      global TM_St_Idle=get_time(STATE_Times[STATE-1])
    elif (5 == switch_1):
      $ 789 "Case 5"
      $ 790 "TM_St_Starting≔get_time(STATE_Times[STATE-1])"
      global TM_St_Starting=get_time(STATE_Times[STATE-1])
    elif (6 == switch_1):
      $ 791 "Case 6"
      $ 792 "TM_St_Execute≔get_time(STATE_Times[STATE-1])"
      global TM_St_Execute=get_time(STATE_Times[STATE-1])
    elif (7 == switch_1):
      $ 793 "Case 7"
      $ 794 "TM_St_Completin≔get_time(STATE_Times[STATE-1])"
      global TM_St_Completin=get_time(STATE_Times[STATE-1])
    elif (8 == switch_1):
      $ 795 "Case 8"
      $ 796 "TM_St_Complete≔get_time(STATE_Times[STATE-1])"
      global TM_St_Complete=get_time(STATE_Times[STATE-1])
    elif (9 == switch_1):
      $ 797 "Case 9"
      $ 798 "TM_St_Holding≔get_time(STATE_Times[STATE-1])"
      global TM_St_Holding=get_time(STATE_Times[STATE-1])
    elif (10 == switch_1):
      $ 799 "Case 10"
      $ 800 "TM_St_Held≔get_time(STATE_Times[STATE-1])"
      global TM_St_Held=get_time(STATE_Times[STATE-1])
    elif (11 == switch_1):
      $ 801 "Case 11"
      $ 802 "TM_St_Unholding≔get_time(STATE_Times[STATE-1])"
      global TM_St_Unholding=get_time(STATE_Times[STATE-1])
    elif (12 == switch_1):
      $ 803 "Case 12"
      $ 804 "TM_St_Suspendin≔get_time(STATE_Times[STATE-1])"
      global TM_St_Suspendin=get_time(STATE_Times[STATE-1])
    elif (13 == switch_1):
      $ 805 "Case 13"
      $ 806 "TM_St_Suspended≔get_time(STATE_Times[STATE-1])"
      global TM_St_Suspended=get_time(STATE_Times[STATE-1])
    elif (14 == switch_1):
      $ 807 "Case 14"
      $ 808 "TM_St_Unsuspend≔get_time(STATE_Times[STATE-1])"
      global TM_St_Unsuspend=get_time(STATE_Times[STATE-1])
    elif (15 == switch_1):
      $ 809 "Case 15"
      $ 810 "TM_St_Aborting≔get_time(STATE_Times[STATE-1])"
      global TM_St_Aborting=get_time(STATE_Times[STATE-1])
    elif (16 == switch_1):
      $ 811 "Case 16"
      $ 812 "TM_St_Aborted≔get_time(STATE_Times[STATE-1])"
      global TM_St_Aborted=get_time(STATE_Times[STATE-1])
    elif (17 == switch_1):
      $ 813 "Case 17"
      $ 814 "TM_St_Clearing≔get_time(STATE_Times[STATE-1])"
      global TM_St_Clearing=get_time(STATE_Times[STATE-1])
    end
    $ 816 "Wait: 0.1"
    sleep(0.1)
  end
end
